ORGANIZATION_BLOCK "Main"
{ S7_Optimized_Access := 'TRUE' }
VERSION : 0.1

BEGIN
	// The standard program only reads what the safety program released.
	"Running" := "SafetyData".released;

END_ORGANIZATION_BLOCK

